Fanuc KAREL source: KT00898.KL

PROGRAM KT00898
%NOLOCKGROUP
VAR
  P1: POSITION
  P2: POSITION
  OUT: BOOLEAN
BEGIN
  OUT = J_IN_RANGE(P1)
END KT00898
